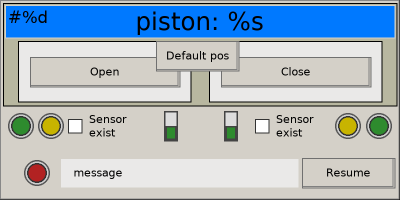
VISUALIZATION vis_Piston_Control1  // 400x200
VAR_IN_OUT
	stPis: ST_Piston;
END_VAR
    Rectangle (0,0 400x200)
    Rectangle (3,3 394x103), colour toggle: NOT stPis.b_Enable
    Rectangle (18,41 173x61), colour toggle: stPis.st_Open
    Rectangle (209,41 173x61), colour toggle: stPis.st_Close
    Button (30,57 150x30), "Open", colour toggle: stPis.req_Open, input disabled if: stPis.b_DeactivateMan OR NOT stPis.b_InterLock_Open
        toggle stPis.req_OpenMan
    Button (221,57 150x30), "Close", colour toggle: stPis.req_Close, input disabled if: stPis.b_DeactivateMan OR NOT stPis.b_InterLock_Close
        toggle stPis.req_CloseMan
    DipSwitch (156,111 30x30), tooltip "Open Sensor state", variable: stPis.sen_Open, invisible if: NOT stPis.sen_Open_Exist, behaviour: TOGGLE, style: Switch-DipSwitch-Green
    DipSwitch (216,111 30x30), tooltip "Close Sensor state", variable: stPis.sen_Close, invisible if: NOT stPis.sen_Close_Exist, behaviour: TOGGLE, style: Switch-DipSwitch-Green
    Checkbox (66,108 99x36), "Sensor exist", variable: stPis.sen_Open_Exist
    Checkbox (253,108 99x36), "Sensor exist", variable: stPis.sen_Close_Exist
    Lamp1 (6,111 30x30), tooltip "Open sensor", variable: stPis.sen_Open, invisible if: NOT stPis.sen_Open_Exist, style: Lamp-Lamp1-Green
    Lamp1 (333,111 30x30), tooltip "Close valve", variable: stPis.valve_Close, style: Lamp-Lamp1-Yellow
    Lamp1 (22,158 30x30), tooltip "Error", variable: stPis.b_Error, style: Lamp-Lamp1-Red
    Textfield (60,158 239x30), "message"
    Button (302,158 93x30), "Resume", colour toggle: stPis.b_Error
        toggle stPis.b_Resume
    Button (156,41 83x30), "Default pos", colour toggle: stPis.req_DefaultPos, input disabled if: stPis.b_DeactivateMan
        toggle stPis.req_DefaultPos
    Textfield (5,5 390x33), "piston: %s", text variable: stPis.sName
    Textfield (5,7 42x21), "#%d", text variable: stPis.iPisNum
    Lamp1 (36,111 30x30), tooltip "Open valve", variable: stPis.valve_Open, style: Lamp-Lamp1-Yellow
    Lamp1 (364,111 30x30), tooltip "Close sensor", variable: stPis.sen_Close, invisible if: NOT stPis.sen_Close_Exist, style: Lamp-Lamp1-Green
END_VISUALIZATION

(* stored: Version 1.1.0.1, ProductVersion 3.1.4024.12
   Visu vis_Piston_Control1: Id {195027a3-d9d1-4238-ae22-7aee00fe3ad8} *)
